FUNCTION_BLOCK F (* Negative C1: the deterministic translator's form, START to RUN to START *)
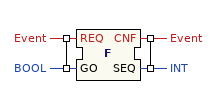
  EVENT_INPUT
    REQ WITH GO;
  END_EVENT
  EVENT_OUTPUT
    CNF WITH SEQ;
  END_EVENT
  VAR_INPUT
    GO : BOOL;
  END_VAR
  VAR_OUTPUT
    SEQ : INT;
  END_VAR
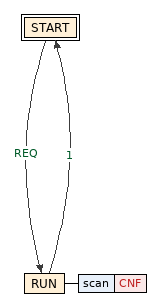
  EC_STATES
    START;
    RUN : scan -> CNF;
  END_STATES
  EC_TRANSITIONS
    START TO RUN := REQ;
    RUN TO START := 1;
  END_TRANSITIONS
  ALGORITHM scan IN ST:
CASE SEQ OF
  0:
    IF GO THEN
      SEQ := 1;
    END_IF;
  1:
    SEQ := 0;
END_CASE;
  END_ALGORITHM
END_FUNCTION_BLOCK
